(* IEC 61131-3 sources: rusty/tests/lit/single/polymorphism, 16 files *)

(* ---- direct_interface_call_does_not_emit_output.st ---- *)
// RUN: rm -f %t.out
// RUN: not %COMPILE --error-format clang %s 2>&1 | %CHECK %s
// RUN: test ! -e %t.out

// Regression test: diagnostics emitted by lowering participants must not produce a binary.
// Lowerers aggregate diagnostics and let the main validation step decide whether to abort,
// so validation errors found during lowering must still stop the pipeline before codegen.

// CHECK: {{.*}}direct_interface_call_does_not_emit_output.st:{{[0-9]+}}:{{[0-9]+}}:{{.*}}error[E129]: Interfaces cannot be called directly
// CHECK: {{.*}}Compilation aborted due to critical errors

INTERFACE IA
    METHOD foo
    END_METHOD
END_INTERFACE

FUNCTION main
    VAR
        refIA : IA;
    END_VAR

    refIA();
END_FUNCTION

(* ---- basic_inheritance.st ---- *)
// RUN: %COMPILE %s && %RUN | %CHECK %s

FUNCTION_BLOCK A
    VAR
        nameA: STRING := 'A';
    END_VAR

    METHOD getName: STRING
        getName := nameA;
    END_METHOD

    METHOD printName
        printf('name = %s$N', ADR(getName()));
    END_METHOD

    METHOD printAncestors
        printf('ancestor = None$N');
    END_METHOD
END_FUNCTION_BLOCK

FUNCTION_BLOCK B EXTENDS A
    VAR
        nameB: STRING := 'B';
    END_VAR

    // OVERRIDE
    METHOD getName: STRING
        getName := nameB;
    END_METHOD

    METHOD printAncestors
        printf('ancestor = %s$N', ADR(SUPER^.getName()));
    END_METHOD
END_FUNCTION_BLOCK

FUNCTION_BLOCK C EXTENDS B
    VAR
        nameC: STRING := 'C';
    END_VAR

    // OVERRIDE
    METHOD getName: STRING
        getName := nameC;
    END_METHOD

    METHOD printAncestors
        SUPER^.printAncestors();
        printf('ancestor = %s$N', ADR(SUPER^.getName()));
    END_METHOD
END_FUNCTION_BLOCK

FUNCTION_BLOCK DD EXTENDS C
    VAR
        nameD: STRING := 'D';
    END_VAR

    // OVERRIDE
    METHOD getName: STRING
        getName := nameD;
    END_METHOD

    METHOD printAncestors
        SUPER^.printAncestors();
        printf('ancestor = %s$N', ADR(SUPER^.getName()));
    END_METHOD
END_FUNCTION_BLOCK

FUNCTION printRefA
    VAR_INPUT
        refInstance: POINTER TO A;
    END_VAR

    refInstance^.printName();
    refInstance^.printAncestors();
END_FUNCTION

FUNCTION main
    VAR
        instanceA: A;
        instanceB: B;
        instanceC: C;
        instanceD: DD;

        refInstanceA: POINTER TO A;
        refInstanceB: POINTER TO B;
        refInstanceC: POINTER TO C;
        refInstanceD: POINTER TO DD;
    END_VAR

    // CHECK: name = A
    // CHECK: ancestor = None
    printRefA(ADR(instanceA));
    printf('$N');

    // CHECK: name = B
    // CHECK: ancestor = A
    printRefA(ADR(instanceB));
    printf('$N');

    // CHECK: name = C
    // CHECK: ancestor = A
    // CHECK: ancestor = B
    printRefA(ADR(instanceC));
    printf('$N');

    // CHECK: name = D
    // CHECK: ancestor = A
    // CHECK: ancestor = B
    // CHECK: ancestor = C
    printRefA(ADR(instanceD));
END_FUNCTION

(* ---- basic_override_method_call_in_method.st ---- *)
// RUN: %COMPILE %s && %RUN | %CHECK %s

FUNCTION_BLOCK A
    VAR
        nameA: STRING := 'A';
    END_VAR

    METHOD getName: STRING
        getName := nameA;
    END_METHOD

    METHOD printName
        printf('name = %s$N', ADR(getName()));
    END_METHOD
END_FUNCTION_BLOCK

FUNCTION_BLOCK B EXTENDS A
    VAR
        nameB: STRING := 'B';
    END_VAR

    // OVERRIDE
    METHOD getName: STRING
        getName := nameB;
    END_METHOD
END_FUNCTION_BLOCK

FUNCTION main
    VAR
        instanceA: A;
        instanceB: B;
        refInstanceA: POINTER TO A;
    END_VAR

    // CHECK: name = A
    refInstanceA := ADR(instanceA);
    refInstanceA^.printName();

    // CHECK: name = B
    refInstanceA := ADR(instanceB);
    refInstanceA^.printName();
END_FUNCTION

(* ---- basic_override_no_method_call_in_method.st ---- *)
// RUN: %COMPILE %s && %RUN | %CHECK %s

FUNCTION_BLOCK A
    METHOD compute : INT
        VAR_INPUT
            value: INT;
        END_VAR

        compute := value * 2;
        printf('A::compute(%d) = %d$N', value, compute);
    END_METHOD
END_FUNCTION_BLOCK

FUNCTION_BLOCK B EXTENDS A
    METHOD compute : INT
        VAR_INPUT
            value: INT;
        END_VAR

        compute := value * 3;
        printf('B::compute(%d) = %d$N', value, compute);
    END_METHOD
END_FUNCTION_BLOCK

FUNCTION processValue : INT
    VAR_INPUT
        obj: POINTER TO A;
        input: INT;
    END_VAR

    processValue := obj^.compute(input);
END_FUNCTION

FUNCTION main
    VAR
        instanceA: A;
        instanceB: B;
        objRef: POINTER TO A;
        result: INT;
    END_VAR

    // ~~ Direct polymorphic calls ~~
    // CHECK: A::compute(5) = 10
    // CHECK: B::compute(5) = 15

    objRef := ADR(instanceA);
    result := objRef^.compute(5);

    objRef := ADR(instanceB);
    result := objRef^.compute(5);

    // ~~ Polymorphic calls through function ~~
    // CHECK: A::compute(7) = 14
    // CHECK: B::compute(7) = 21

    objRef := ADR(instanceA);
    result := processValue(objRef, 7);

    objRef := ADR(instanceB);
    result := processValue(objRef, 7);
END_FUNCTION

(* ---- calls_through_pointer_in_method.st ---- *)
// RUN: %COMPILE %s && %RUN | %CHECK %s
// Scenario: A method or body of one POU calls methods and properties of another function block through a
// `REFERENCE TO` or a `POINTER TO`. The call must dispatch through the virtual table of that instance, not
// of the enclosing POU, also when the enclosing POU has a method with the same name. This holds in function
// blocks, classes, and programs, and a derived instance behind the pointer runs its override. A body call
// through a qualified reference, `refBox.target()`, uses the type of `target`, not of `refBox`.

TYPE Box : STRUCT
    target : REFERENCE TO fb;
END_STRUCT END_TYPE

FUNCTION_BLOCK fb
    VAR
        stored : INT;
        bodyCalls : DINT;
    END_VAR

    PROPERTY_GET prop : INT
        prop := stored;
    END_PROPERTY

    PROPERTY_SET prop : INT
        stored := prop;
    END_PROPERTY

    METHOD foo : DINT
        foo := 42;
    END_METHOD

    METHOD add : DINT
        VAR_INPUT
            a : DINT;
        END_VAR

        add := a + 100;
    END_METHOD

    bodyCalls := bodyCalls + 1;
END_FUNCTION_BLOCK

FUNCTION_BLOCK fbDerived EXTENDS fb
    METHOD foo : DINT
        foo := 43;
    END_METHOD
END_FUNCTION_BLOCK

FUNCTION_BLOCK holder
    VAR
        rfb : REFERENCE TO fb;
        pfb : POINTER TO fb;
        refBox : REFERENCE TO Box;
        bodyResult : DINT;
    END_VAR

    METHOD a : DINT
        a := 1;
    END_METHOD

    METHOD foo : DINT
        foo := 3;
    END_METHOD

    METHOD run : DINT
        rfb.prop := rfb.prop + 1;
        pfb^.prop := pfb^.prop + 1;
        run := rfb.foo() * 1000 + pfb^.add(5) + foo();
    END_METHOD

    METHOD runTarget
        refBox.target();
    END_METHOD

    bodyResult := pfb^.foo();
END_FUNCTION_BLOCK

CLASS user
    VAR
        pfb : POINTER TO fb;
    END_VAR

    METHOD foo : DINT
        foo := 4;
    END_METHOD

    METHOD run : DINT
        run := pfb^.foo();
    END_METHOD
END_CLASS

PROGRAM mainProg
    VAR
        myfb : fb;
        rfb : REFERENCE TO fb;
        pfb : POINTER TO fb;
    END_VAR

    METHOD baz : INT
        myfb.prop := myfb.prop + 1;
        myfb.foo();

        rfb.prop := rfb.prop + 1;
        rfb.foo();

        pfb^.prop := pfb^.prop + 1;
        pfb^.foo();

        baz := myfb.prop;
    END_METHOD
END_PROGRAM

FUNCTION runTargetFromFunction
    VAR_INPUT
        ptrBox : REF_TO Box;
    END_VAR
    VAR
        rbox : REFERENCE TO Box;
    END_VAR

    rbox REF= ptrBox^;
    rbox.target();
END_FUNCTION

FUNCTION main : DINT
    VAR
        f : fb;
        d : fbDerived;
        h : holder;
        u : user;
        b : Box;
    END_VAR

    // CHECK: holder: 42108 2
    h.rfb REF= f;
    h.pfb := ADR(f);
    printf('holder: %d %d$N', h.run(), f.prop);

    // CHECK: holder body: 43
    h.pfb := ADR(d);
    h();
    printf('holder body: %d$N', h.bodyResult);

    // CHECK: class: 43
    u.pfb := ADR(d);
    printf('class: %d$N', u.run());

    // CHECK: body through qualified reference: 2
    b.target REF= f;
    h.refBox REF= b;
    h.runTarget();
    runTargetFromFunction(REF(b));
    printf('body through qualified reference: %d$N', f.bodyCalls);

    // CHECK: program: 3
    mainProg.rfb REF= mainProg.myfb;
    mainProg.pfb := ADR(mainProg.myfb);
    printf('program: %d$N', mainProg.baz());
END_FUNCTION

(* ---- function_block_call.st ---- *)
// RUN: %COMPILE %s && %RUN | %CHECK %s

FUNCTION_BLOCK A
    VAR
        localStateA: DINT := 1;
    END_VAR

    printf('A::body: localStateA = %d$N', localStateA);
END_FUNCTION_BLOCK

FUNCTION_BLOCK B EXTENDS A
    VAR
        localStateB: DINT := 2;
    END_VAR

    SUPER^();
    printf('B::body: localStateB = %d$N', localStateB);
END_FUNCTION_BLOCK

FUNCTION_BLOCK C EXTENDS B
    VAR
        localStateC: DINT := 3;
    END_VAR

    SUPER^();
    printf('C::body: localStateC = %d$N', localStateC);
END_FUNCTION_BLOCK

FUNCTION main
    VAR
        instanceA: A;
        instanceB: B;
        instanceC: C;

        refInstanceA: POINTER TO A;
        refInstanceB: POINTER TO B;
        refInstanceC: POINTER TO C;
    END_VAR

    instanceA.localStateA := 5;
    instanceB.localStateB := 10;
    instanceC.localStateC := 15;

    // CHECK: A::body: localStateA = 5
    refInstanceA := ADR(instanceA);
    refInstanceA^();

    // CHECK: A::body: localStateA = 1
    // CHECK: B::body: localStateB = 10
    refInstanceA := ADR(instanceB);
    refInstanceA^();

    // CHECK: A::body: localStateA = 1
    // CHECK: B::body: localStateB = 2
    // CHECK: C::body: localStateC = 15
    refInstanceA := ADR(instanceC);
    refInstanceA^();

    // CHECK: A::body: localStateA = 1
    // CHECK: B::body: localStateB = 10
    refInstanceB := ADR(instanceB);
    refInstanceB^();

    // CHECK: A::body: localStateA = 1
    // CHECK: B::body: localStateB = 2
    // CHECK: C::body: localStateC = 15
    refInstanceB := ADR(instanceC);
    refInstanceB^();

    // CHECK: A::body: localStateA = 1
    // CHECK: B::body: localStateB = 2
    // CHECK: C::body: localStateC = 15
    refInstanceC := ADR(instanceC);
    refInstanceC^();
END_FUNCTION

(* ---- inheritance_chain.st ---- *)
// RUN: %COMPILE %s && %RUN | %CHECK %s

FUNCTION_BLOCK A
    METHOD printName: STRING
        printf('FB A$N');
    END_METHOD

    METHOD A1
        printf('  A::A1$N');
    END_METHOD

    METHOD A2
        printf('  A::A2$N');
    END_METHOD

    METHOD A3
        printf('  A::A3$N');
    END_METHOD

    METHOD A4
        printf('  A::A4$N');
    END_METHOD

    METHOD callMethods
        A1();
        A2();
        A3();
        A4();
    END_METHOD
END_FUNCTION_BLOCK

// B overriddes A2, introduces B1, B2 and B3
FUNCTION_BLOCK B EXTENDS A
    METHOD printName: STRING
        printf('FB B$N');
    END_METHOD

    METHOD A2
        printf('  B::A2 (overridden)$N');
    END_METHOD

    METHOD B1
        printf('  B::B1$N');
    END_METHOD

    METHOD B2
        printf('  B::B2$N');
    END_METHOD

    METHOD B3
        printf('  B::B3$N');
    END_METHOD
END_FUNCTION_BLOCK

// C overriddes A3, B2, introduces C1 and C2
FUNCTION_BLOCK C EXTENDS B
    METHOD printName: STRING
        printf('FB C$N');
    END_METHOD

    METHOD A3
        printf('  C::A3 (overridden)$N');
    END_METHOD

    METHOD B2
        printf('  C::B2 (overridden)$N');
    END_METHOD

    METHOD C1
        printf('  C::C1$N');
    END_METHOD

    METHOD C2
        printf('  C::C2$N');
    END_METHOD
END_FUNCTION_BLOCK

// D overriddes A4, B3, C2, introduces D1
FUNCTION_BLOCK DD EXTENDS C
    METHOD printName: STRING
        printf('FB D$N');
    END_METHOD

    METHOD A4
        printf('  D::A4 (overridden)$N');
    END_METHOD

    METHOD B3
        printf('  D::B3 (overridden)$N');
    END_METHOD

    METHOD C2
        printf('  D::C2 (overridden)$N');
    END_METHOD

    METHOD D1
        printf('  D::D1$N');
    END_METHOD
END_FUNCTION_BLOCK

FUNCTION main
    VAR
        index: INT;

        instanceA: A;
        instanceB: B;
        instanceC: C;
        instanceD: DD;

        instanceRefArrayA: ARRAY[1..4] OF POINTER TO A;
        instanceRefArrayB: ARRAY[1..3] OF POINTER TO B;
        instanceRefArrayC: ARRAY[1..2] OF POINTER TO C;
        instanceRefArrayD: ARRAY[1..1] OF POINTER TO DD;
    END_VAR

    // TODOs
    // - initializer in variable declaration not working, e.g. `instanceRefArrayD: ARRAY[1..1] OF POINTER TO D := [ADR(instanceD)]`
    // - initializer in body not working, e.g. `instanceRefArrayD := [ADR(instanceD)]`

    // Initialize the arrays
    instanceRefArrayA[1] := ADR(instanceA);
    instanceRefArrayA[2] := ADR(instanceB);
    instanceRefArrayA[3] := ADR(instanceC);
    instanceRefArrayA[4] := ADR(instanceD);

    instanceRefArrayB[1] := ADR(instanceB);
    instanceRefArrayB[2] := ADR(instanceC);
    instanceRefArrayB[3] := ADR(instanceD);

    instanceRefArrayC[1] := ADR(instanceC);
    instanceRefArrayC[2] := ADR(instanceD);

    instanceRefArrayD[1] := ADR(instanceD);

    // CHECK: -- FUNCTION_BLOCK A and its children --
    // CHECK: FB A
    // CHECK:   A::A1
    // CHECK:   A::A2
    // CHECK:   A::A3
    // CHECK:   A::A4
    // CHECK: FB B
    // CHECK:   A::A1
    // CHECK:   B::A2 (overridden)
    // CHECK:   A::A3
    // CHECK:   A::A4
    // CHECK: FB C
    // CHECK:   A::A1
    // CHECK:   B::A2 (overridden)
    // CHECK:   C::A3 (overridden)
    // CHECK:   A::A4
    // CHECK: FB D
    // CHECK:   A::A1
    // CHECK:   B::A2 (overridden)
    // CHECK:   C::A3 (overridden)
    // CHECK:   D::A4 (overridden)
    printf('-- FUNCTION_BLOCK A and its children --$N');
    FOR index := 1 TO 4 DO
        instanceRefArrayA[index]^.printName();
        instanceRefArrayA[index]^.A1();
        instanceRefArrayA[index]^.A2();
        instanceRefArrayA[index]^.A3();
        instanceRefArrayA[index]^.A4();
    END_FOR

    // CHECK: -- FUNCTION_BLOCK B and its children --
    // CHECK: FB B
    // CHECK:   A::A1
    // CHECK:   B::A2 (overridden)
    // CHECK:   A::A3
    // CHECK:   A::A4
    // CHECK:   B::B1
    // CHECK:   B::B2
    // CHECK:   B::B3
    // CHECK: FB C
    // CHECK:   A::A1
    // CHECK:   B::A2 (overridden)
    // CHECK:   C::A3 (overridden)
    // CHECK:   A::A4
    // CHECK:   B::B1
    // CHECK:   C::B2 (overridden)
    // CHECK:   B::B3
    // CHECK: FB D
    // CHECK:   A::A1
    // CHECK:   B::A2 (overridden)
    // CHECK:   C::A3 (overridden)
    // CHECK:   D::A4 (overridden)
    // CHECK:   B::B1
    // CHECK:   C::B2 (overridden)
    // CHECK:   D::B3 (overridden)
    printf('$N$N-- FUNCTION_BLOCK B and its children --$N');
    FOR index := 1 TO 3 DO
        instanceRefArrayB[index]^.printName();
        instanceRefArrayB[index]^.A1();
        instanceRefArrayB[index]^.A2();
        instanceRefArrayB[index]^.A3();
        instanceRefArrayB[index]^.A4();
        instanceRefArrayB[index]^.B1();
        instanceRefArrayB[index]^.B2();
        instanceRefArrayB[index]^.B3();
    END_FOR

    // CHECK: -- FUNCTION_BLOCK C and its children --
    // CHECK: FB C
    // CHECK:   A::A1
    // CHECK:   B::A2 (overridden)
    // CHECK:   C::A3 (overridden)
    // CHECK:   A::A4
    // CHECK:   B::B1
    // CHECK:   C::B2 (overridden)
    // CHECK:   B::B3
    // CHECK:   C::C1
    // CHECK:   C::C2
    // CHECK: FB D
    // CHECK:   A::A1
    // CHECK:   B::A2 (overridden)
    // CHECK:   C::A3 (overridden)
    // CHECK:   D::A4 (overridden)
    // CHECK:   B::B1
    // CHECK:   C::B2 (overridden)
    // CHECK:   D::B3 (overridden)
    // CHECK:   C::C1
    // CHECK:   D::C2 (overridden)
    printf('$N$N-- FUNCTION_BLOCK C and its children --$N');
    FOR index := 1 TO 2 DO
        instanceRefArrayC[index]^.printName();
        instanceRefArrayC[index]^.A1();
        instanceRefArrayC[index]^.A2();
        instanceRefArrayC[index]^.A3();
        instanceRefArrayC[index]^.A4();
        instanceRefArrayC[index]^.B1();
        instanceRefArrayC[index]^.B2();
        instanceRefArrayC[index]^.B3();
        instanceRefArrayC[index]^.C1();
        instanceRefArrayC[index]^.C2();
    END_FOR

    // CHECK: -- FUNCTION_BLOCK D and its children (it doesnt have any 😔) --
    // CHECK: FB D
    // CHECK:   A::A1
    // CHECK:   B::A2 (overridden)
    // CHECK:   C::A3 (overridden)
    // CHECK:   D::A4 (overridden)
    // CHECK:   B::B1
    // CHECK:   C::B2 (overridden)
    // CHECK:   D::B3 (overridden)
    // CHECK:   C::C1
    // CHECK:   D::C2 (overridden)
    // CHECK:   D::D1
    printf('$N$N-- FUNCTION_BLOCK D and its children (it doesnt have any 😔) --$N');
    FOR index := 1 TO 1 DO
        instanceRefArrayD[index]^.printName();
        instanceRefArrayD[index]^.A1();
        instanceRefArrayD[index]^.A2();
        instanceRefArrayD[index]^.A3();
        instanceRefArrayD[index]^.A4();
        instanceRefArrayD[index]^.B1();
        instanceRefArrayD[index]^.B2();
        instanceRefArrayD[index]^.B3();
        instanceRefArrayD[index]^.C1();
        instanceRefArrayD[index]^.C2();
        instanceRefArrayD[index]^.D1();
    END_FOR
END_FUNCTION

(* ---- pointer_call_in_function_block.st ---- *)
// RUN: %COMPILE %s && %RUN | %CHECK %s

FUNCTION_BLOCK A
    VAR_INPUT
        in: DINT;
    END_VAR

    METHOD alpha: DINT
        alpha := 1;
    END_METHOD

    METHOD compute: DINT
        compute := 2;
    END_METHOD

    printf('A body, in = %d$N', in);
END_FUNCTION_BLOCK

FUNCTION_BLOCK B EXTENDS A
    METHOD compute: DINT
        compute := 3;
    END_METHOD

    printf('B body, in = %d$N', in);
END_FUNCTION_BLOCK

// `compute` of C is in a different vtable slot than `compute` of A
FUNCTION_BLOCK C
    VAR_INPUT
        refToA: REF_TO A;
        pointerToA: POINTER TO A;
        referenceToA: REFERENCE TO A;
    END_VAR

    METHOD compute: DINT
        compute := 99;
    END_METHOD

    METHOD printFromMethod
        printf('method: ref_to = %d, pointer_to = %d, reference_to = %d$N', refToA^.compute(), pointerToA^.compute(), referenceToA.compute());
    END_METHOD

    printf('body: ref_to = %d, pointer_to = %d, reference_to = %d$N', refToA^.compute(), pointerToA^.compute(), referenceToA.compute());
    referenceToA(in := 7);
END_FUNCTION_BLOCK

CLASS Reader
    VAR
        refToA: REF_TO A;
    END_VAR

    METHOD printFromClass
        VAR_INPUT
            target: REF_TO A;
        END_VAR

        refToA := target;
        printf('class: ref_to = %d$N', refToA^.compute());
    END_METHOD
END_CLASS

FUNCTION main
    VAR
        instanceA: A;
        instanceB: B;
        instanceC: C;
        instanceReader: Reader;
    END_VAR

    // CHECK: body: ref_to = 2, pointer_to = 2, reference_to = 2
    // CHECK: A body, in = 7
    // CHECK: method: ref_to = 2, pointer_to = 2, reference_to = 2
    instanceC.referenceToA REF= instanceA;
    instanceC(refToA := REF(instanceA), pointerToA := ADR(instanceA));
    instanceC.printFromMethod();

    // CHECK: body: ref_to = 3, pointer_to = 3, reference_to = 3
    // CHECK: B body, in = 7
    // CHECK: method: ref_to = 3, pointer_to = 3, reference_to = 3
    instanceC.referenceToA REF= instanceB;
    instanceC(refToA := REF(instanceB), pointerToA := ADR(instanceB));
    instanceC.printFromMethod();

    // CHECK: class: ref_to = 2
    // CHECK: class: ref_to = 3
    instanceReader.printFromClass(REF(instanceA));
    instanceReader.printFromClass(REF(instanceB));
END_FUNCTION

(* ---- pointer_to_pointer_upcast.st ---- *)
// RUN: %COMPILE %s && %RUN | %CHECK %s

FUNCTION_BLOCK A
    METHOD getName: STRING
        getName := 'A';
    END_METHOD
END_FUNCTION_BLOCK

FUNCTION_BLOCK B EXTENDS A
    METHOD getName: STRING
        getName := 'B';
    END_METHOD
END_FUNCTION_BLOCK

FUNCTION_BLOCK C EXTENDS B
    METHOD getName: STRING
        getName := 'C';
    END_METHOD
END_FUNCTION_BLOCK

FUNCTION main
    VAR
        instanceA: A;
        instanceB: B;
        instanceC: C;

        ptrA: POINTER TO A;
        ptrB: POINTER TO B;
        ptrC: POINTER TO C;
    END_VAR

    // Pointer-to-pointer upcast: assign child pointer to base pointer
    ptrB := ADR(instanceB);
    ptrA := ptrB;
    // CHECK: name = B
    printf('name = %s$N', ADR(ptrA^.getName()));

    ptrC := ADR(instanceC);
    ptrA := ptrC;
    // CHECK: name = C
    printf('name = %s$N', ADR(ptrA^.getName()));

    // Transitive: ptrC -> ptrB -> ptrA
    ptrC := ADR(instanceC);
    ptrB := ptrC;
    ptrA := ptrB;
    // CHECK: name = C
    printf('name = %s$N', ADR(ptrA^.getName()));
END_FUNCTION

(* ---- property_vtable_dispatch.st ---- *)
// RUN: %COMPILE %s && %RUN | %CHECK %s
// Scenario: POU-based polymorphism (vtable dispatch) with properties. A method in the base FB
// accesses a property. When the property getter is overridden in a child FB, calling that method
// through a pointer-to-base should dispatch to the overridden getter via the vtable.

FUNCTION_BLOCK A
    VAR
        _val : DINT := 10;
    END_VAR

    PROPERTY_GET value: DINT
        value := _val;
    END_PROPERTY

    PROPERTY_SET value: DINT
        _val := value;
    END_PROPERTY

    METHOD printValue
        printf('value=%d$N', value);
    END_METHOD

    METHOD setValue
        VAR_INPUT x : DINT; END_VAR
        value := x;
    END_METHOD
END_FUNCTION_BLOCK

FUNCTION_BLOCK B EXTENDS A
    // Override getter — adds 1000 to distinguish from A's getter
    PROPERTY_GET value: DINT
        value := _val + 1000;
    END_PROPERTY
END_FUNCTION_BLOCK

FUNCTION_BLOCK C EXTENDS B
    // Override getter again — adds 2000
    PROPERTY_GET value: DINT
        value := _val + 2000;
    END_PROPERTY
END_FUNCTION_BLOCK

FUNCTION printViaPtr
    VAR_INPUT
        refInstance : POINTER TO A;
    END_VAR

    refInstance^.printValue();
END_FUNCTION

FUNCTION setViaPtr
    VAR_INPUT
        refInstance : POINTER TO A;
        x : DINT;
    END_VAR

    refInstance^.setValue(x);
END_FUNCTION

FUNCTION setDirectViaPtr
    VAR_INPUT
        refInstance : POINTER TO A;
        x : DINT;
    END_VAR

    refInstance^.value := x;
END_FUNCTION

FUNCTION main
    VAR
        instanceA : A;
        instanceB : B;
        instanceC : C;
    END_VAR

    // A — base getter
    printViaPtr(ADR(instanceA));        // CHECK: value=10

    // B — overridden getter adds 1000
    printViaPtr(ADR(instanceB));        // CHECK-NEXT: value=1010

    // C — overridden getter adds 2000
    printViaPtr(ADR(instanceC));        // CHECK-NEXT: value=2010

    // Setter through pointer on B (inherited from A), then read with overridden getter
    setViaPtr(ADR(instanceB), 42);
    printViaPtr(ADR(instanceB));        // CHECK-NEXT: value=1042

    // Setter through pointer on C, then read with C's getter
    setViaPtr(ADR(instanceC), 99);
    printViaPtr(ADR(instanceC));        // CHECK-NEXT: value=2099

    // Direct access on concrete instances still works
    printf('value=%d$N', instanceA.value);  // CHECK-NEXT: value=10
    printf('value=%d$N', instanceB.value);  // CHECK-NEXT: value=1042
    printf('value=%d$N', instanceC.value);  // CHECK-NEXT: value=2099

    // Direct property setter through pointer (not via method)
    setDirectViaPtr(ADR(instanceA), 77);
    printViaPtr(ADR(instanceA));            // CHECK-NEXT: value=77

    setDirectViaPtr(ADR(instanceB), 55);
    printViaPtr(ADR(instanceB));            // CHECK-NEXT: value=1055

    setDirectViaPtr(ADR(instanceC), 33);
    printViaPtr(ADR(instanceC));            // CHECK-NEXT: value=2033
END_FUNCTION

(* ---- ref_to.st ---- *)
// RUN: %COMPILE %s && %RUN | %CHECK %s

FUNCTION_BLOCK A
    METHOD alpha
        printf('A::alpha$N');
    END_METHOD

    METHOD bravo
        printf('A::bravo$N');
    END_METHOD

    printf('A::body$N');
END_FUNCTION_BLOCK

FUNCTION_BLOCK B EXTENDS A
    METHOD alpha
        printf('B::alpha$N');
    END_METHOD

    printf('B::body$N');
END_FUNCTION_BLOCK

FUNCTION_BLOCK C EXTENDS B
    METHOD alpha
        printf('C::alpha$N');
    END_METHOD

    METHOD bravo
        printf('C::bravo$N');
    END_METHOD

    printf('C::body$N');
END_FUNCTION_BLOCK

FUNCTION main
    VAR
        instanceA: A;
        instanceB: B;
        instanceC: C;

        refInstanceA: REF_TO A;
    END_VAR

    // CHECK: A::body
    // CHECK: A::alpha
    // CHECK: A::bravo
    refInstanceA := REF(instanceA);
    refInstanceA^();
    refInstanceA^.alpha();
    refInstanceA^.bravo();

    // CHECK: B::body
    // CHECK: B::alpha
    // CHECK: A::bravo
    refInstanceA := REF(instanceB);
    refInstanceA^();
    refInstanceA^.alpha();
    refInstanceA^.bravo();

    // CHECK: C::body
    // CHECK: C::alpha
    // CHECK: C::bravo
    refInstanceA := REF(instanceC);
    refInstanceA^();
    refInstanceA^.alpha();
    refInstanceA^.bravo();
END_FUNCTION

(* ---- reference_to.st ---- *)
// RUN: %COMPILE %s && %RUN | %CHECK %s

FUNCTION_BLOCK A
    METHOD alpha
        printf('A::alpha$N');
    END_METHOD

    METHOD bravo
        printf('A::bravo$N');
    END_METHOD

    printf('A::body$N');
END_FUNCTION_BLOCK

FUNCTION_BLOCK B EXTENDS A
    METHOD alpha
        printf('B::alpha$N');
    END_METHOD

    printf('B::body$N');
END_FUNCTION_BLOCK

FUNCTION_BLOCK C EXTENDS B
    METHOD alpha
        printf('C::alpha$N');
    END_METHOD

    METHOD bravo
        printf('C::bravo$N');
    END_METHOD

    printf('C::body$N');
END_FUNCTION_BLOCK

FUNCTION main
    VAR
        instanceA: A;
        instanceB: B;
        instanceC: C;

        refInstanceA: REFERENCE TO A;
    END_VAR

    // CHECK: A::body
    // CHECK: A::alpha
    // CHECK: A::bravo
    refInstanceA REF= instanceA;
    refInstanceA();
    refInstanceA.alpha();
    refInstanceA.bravo();

    // CHECK: B::body
    // CHECK: B::alpha
    // CHECK: A::bravo
    refInstanceA REF= instanceB;
    refInstanceA();
    refInstanceA.alpha();
    refInstanceA.bravo();

    // CHECK: C::body
    // CHECK: C::alpha
    // CHECK: C::bravo
    refInstanceA REF= instanceC;
    refInstanceA();
    refInstanceA.alpha();
    refInstanceA.bravo();
END_FUNCTION

(* ---- super_call.st ---- *)
// RUN: %COMPILE %s && %RUN | %CHECK %s

FUNCTION_BLOCK A
    METHOD foo
        printf('A::foo$N');
    END_METHOD

    printf('A::body$N');
END_FUNCTION_BLOCK

FUNCTION_BLOCK B EXTENDS A
    METHOD foo
        printf('B::foo$N');
        SUPER^.foo();
        SUPER^();
    END_METHOD

    printf('B::body$N');
END_FUNCTION_BLOCK

FUNCTION_BLOCK C EXTENDS B
    METHOD foo
        printf('C::foo$N');
        SUPER^.foo();
        SUPER^();
    END_METHOD

    printf('C::body$N');
END_FUNCTION_BLOCK

FUNCTION main
    VAR
        instanceA: A;
        instanceB: B;
        instanceC: C;

        refInstanceA: POINTER TO A;
    END_VAR

    // CHECK: A::foo
    refInstanceA := ADR(instanceA);
    refInstanceA^.foo();

    // CHECK: B::foo
    // CHECK: A::foo
    // CHECK: A::body
    refInstanceA := ADR(instanceB);
    refInstanceA^.foo();

    // CHECK: C::foo
    // CHECK: B::foo
    // CHECK: A::foo
    // CHECK: A::body
    // CHECK: B::body
    refInstanceA := ADR(instanceC);
    refInstanceA^.foo();
END_FUNCTION

(* ---- this_call.st ---- *)
// RUN: %COMPILE %s && %RUN | %CHECK %s

FUNCTION_BLOCK A
    METHOD foo
        printf('A::foo$N');
        THIS^();
    END_METHOD

    printf('A::body$N');
END_FUNCTION_BLOCK

FUNCTION_BLOCK B EXTENDS A
    METHOD bar
        THIS^();
    END_METHOD

    printf('B::body$N');
END_FUNCTION_BLOCK

FUNCTION_BLOCK C EXTENDS B
    METHOD foo
        printf('C::foo$N');
        THIS^();
    END_METHOD

    printf('C::body$N');
END_FUNCTION_BLOCK

FUNCTION main
    VAR
        instanceA: A;
        instanceB: B;
        instanceC: C;

        refInstanceA: POINTER TO A;
    END_VAR

    // CHECK: A::foo
    // CHECK: A::body
    refInstanceA := ADR(instanceA);
    refInstanceA^.foo();

    // CHECK: A::foo
    // CHECK: A::body
    refInstanceA := ADR(instanceB);
    refInstanceA^.foo();

    // CHECK: C::foo
    // CHECK: C::body
    refInstanceA := ADR(instanceC);
    refInstanceA^.foo();
END_FUNCTION

(* ---- this_method_call.st ---- *)
// RUN: %COMPILE %s && %RUN | %CHECK %s
// Scenario: `THIS^.foo()` stands for the actual instance, so it dispatches through the vtable exactly
// like the unqualified `foo()`. A child or grandchild override must run, also for property accessors,
// for calls with named arguments and outputs, and for the body of a base that a child runs via `SUPER^()`.

FUNCTION_BLOCK Dog
    VAR
        bodyResult : DINT;
        stored : DINT;
    END_VAR

    METHOD say : DINT
        say := 1;
    END_METHOD

    METHOD add : DINT
        VAR_INPUT
            a : DINT;
        END_VAR
        VAR_OUTPUT
            tag : DINT;
        END_VAR

        add := a + 10;
        tag := 1;
    END_METHOD

    PROPERTY_GET name : DINT
        name := 1;
    END_PROPERTY

    PROPERTY_SET level : DINT
        stored := level;
    END_PROPERTY

    METHOD plain : DINT
        plain := say();
    END_METHOD

    METHOD viaThis : DINT
        viaThis := THIS^.say();
    END_METHOD

    METHOD viaThisNamed : DINT
        VAR
            t : DINT;
        END_VAR

        viaThisNamed := THIS^.add(a := 5, tag => t) * 10 + t;
    END_METHOD

    METHOD viaThisProperty : DINT
        viaThisProperty := THIS^.name;
    END_METHOD

    METHOD setViaThis
        THIS^.level := 7;
    END_METHOD

    bodyResult := THIS^.say();
END_FUNCTION_BLOCK

FUNCTION_BLOCK Puppy EXTENDS Dog
    METHOD say : DINT
        say := 2;
    END_METHOD

    METHOD add : DINT
        VAR_INPUT
            a : DINT;
        END_VAR
        VAR_OUTPUT
            tag : DINT;
        END_VAR

        add := a + 20;
        tag := 2;
    END_METHOD

    PROPERTY_GET name : DINT
        name := 2;
    END_PROPERTY

    PROPERTY_SET level : DINT
        stored := level * 100;
    END_PROPERTY

    SUPER^();
END_FUNCTION_BLOCK

FUNCTION_BLOCK Pup EXTENDS Puppy
    METHOD say : DINT
        say := 3;
    END_METHOD

    SUPER^();
END_FUNCTION_BLOCK

FUNCTION main : DINT
    VAR
        d : Dog;
        p : Puppy;
        g : Pup;
        ref : POINTER TO Dog;
    END_VAR

    // CHECK: plain: 1 2 3
    printf('plain: %d %d %d$N', d.plain(), p.plain(), g.plain());

    // CHECK: viaThis: 1 2 3
    printf('viaThis: %d %d %d$N', d.viaThis(), p.viaThis(), g.viaThis());

    // CHECK: viaThisNamed: 151 252 252
    printf('viaThisNamed: %d %d %d$N', d.viaThisNamed(), p.viaThisNamed(), g.viaThisNamed());

    // CHECK: viaThisProperty: 1 2 2
    printf('viaThisProperty: %d %d %d$N', d.viaThisProperty(), p.viaThisProperty(), g.viaThisProperty());

    // CHECK: setViaThis: 7 700 700
    d.setViaThis();
    p.setViaThis();
    g.setViaThis();
    printf('setViaThis: %d %d %d$N', d.stored, p.stored, g.stored);

    // CHECK: viaPointer: 3
    ref := ADR(g);
    printf('viaPointer: %d$N', ref^.viaThis());

    // CHECK: body: 1 2 3
    d();
    p();
    g();
    printf('body: %d %d %d$N', d.bodyResult, p.bodyResult, g.bodyResult);
END_FUNCTION

(* ---- unordered_method_declaration.st ---- *)
// RUN: %COMPILE %s && %RUN | %CHECK %s
// This test ensures that even with an unordered method declaration, the methods internally are still defined
// in a fixed order within the virtual table. Specifically, if function block A defines methods in order
// [alpha, bravo, charlie] and function block B extends A overridding bravo and introducing delta in order
// [delta, bravo] then internally the virtual table must be defined as [alpha, bravo, charlie, delta] rather
// than [delta, bravo, alpha, charlie]. Not doing so would break the ability to upcast from B to A because
// B's virtual table would not match the expected layout of its super class A = [alpha, bravo, charlie].

FUNCTION_BLOCK A
    METHOD alpha
        printf('A::alpha$N');
    END_METHOD

    METHOD bravo
        printf('A::bravo$N');
    END_METHOD

    METHOD charlie
        printf('A::charlie$N');
    END_METHOD

    METHOD delta
        printf('A::delta$N');
    END_METHOD

    printf('A::body$N');
END_FUNCTION_BLOCK

FUNCTION_BLOCK B EXTENDS A
    METHOD echo
        printf('B::echo$N');
    END_METHOD

    // Overridden
    METHOD charlie
        printf('B::charlie$N');
    END_METHOD

    // Overridden
    METHOD alpha
        printf('B::alpha$N');
    END_METHOD

    METHOD foxtrot
        printf('B::foxtrot$N');
    END_METHOD

    printf('B::body$N');
END_FUNCTION_BLOCK

FUNCTION_BLOCK C EXTENDS B
    METHOD golf
        printf('C::golf$N');
    END_METHOD

    printf('C::body$N');
END_FUNCTION_BLOCK

FUNCTION main
    VAR
        instanceA: A;
        instanceB: B;
        instanceC: C;

        refInstanceA: POINTER TO A;
    END_VAR

    // CHECK: A::body
    // CHECK: A::alpha
    // CHECK: A::bravo
    // CHECK: A::charlie
    // CHECK: A::delta
    refInstanceA := ADR(instanceA);
    refInstanceA^();
    refInstanceA^.alpha();
    refInstanceA^.bravo();
    refInstanceA^.charlie();
    refInstanceA^.delta();

    // CHECK: B::body
    // CHECK: B::alpha
    // CHECK: A::bravo
    // CHECK: B::charlie
    // CHECK: A::delta
    refInstanceA := ADR(instanceB);
    refInstanceA^();
    refInstanceA^.alpha();
    refInstanceA^.bravo();
    refInstanceA^.charlie();
    refInstanceA^.delta();

    // CHECK: C::body
    // CHECK: B::alpha
    // CHECK: A::bravo
    // CHECK: B::charlie
    // CHECK: A::delta
    refInstanceA := ADR(instanceC);
    refInstanceA^();
    refInstanceA^.alpha();
    refInstanceA^.bravo();
    refInstanceA^.charlie();
    refInstanceA^.delta();
END_FUNCTION
